(* IEC 61131-3 sources: codesys-framework/txt/application/WeVe General (library)/EmergencyStop/DUT, 1 file *)

(* ---- E_EmergencyStopState.dut.st ---- *)
{attribute 'qualified_only'}
{attribute 'strict'}
TYPE E_EmergencyStopState :
(
	OK := 0,
	NOK
);
END_TYPE
